// TIA Portal project "LaboratorioPID" (V21)

(* hardware
DEVICE "S7-1200 station_1"  S7-1200 Station
   slot 0: "Rack_0"  S7-1200 Rack  Rack  V1.0
   slot 1: "PLC-Serrato"  CPU 1214C AC/DC/Rly  6ES7 214-1BG40-0XB0  V4.2
   slot 3: "AQ 1x12BIT_1"  AQ1 signal board  6ES7 232-4HA30-0XB0  V1.0
DEVICE "HMI_1"  TP1200 Comfort
   slot 0: "HMI_1"  TP1200 Comfort  6AV2 124-0MC01-0AX0  17.0.0.0
   slot 1: "HMI_RT_1"  TP1200 Comfort  6AV2 124-0MC01-0AX0  17.0.0.0
   slot 5: "HMI_1.IE_CP_1"  PROFINET Interface  17.0.0.0
      slot 1: "PROFINET Interface_1"  PROFINET Interface
         slot 1: "Port_1"  Port
         slot 2: "Port_2"  Port
   slot 7: "HMI_1.MPI/DP_CP_1"  MPI/DP Interface  17.0.0.0
DEVICE "S7-1200 station_2"  S7-1200 Station
   slot 0: "Rack_0"  S7-1200 Rack  Rack  V1.0
   slot 1: "PLC-Liceth"  CPU 1214C AC/DC/Rly  6ES7 214-1BG40-0XB0  V4.2
*)

// ===== PLC "PLC-Serrato"  CPU 1214C AC/DC/Rly =====

VAR_GLOBAL   // PLC tag table "Default tag table"
   "PresionRaw" AT %IW64 : Int;
   "BelimoRaw" AT %QW80 : Int;
   "PID_salida_pct" AT %MD0 : Real;
   "Apertura_Manual" AT %MD10 : Real;
   "Clock_Byte" AT %MB100 : Byte;
   "Clock_10Hz" AT %M100.0 : Bool;
   "Clock_5Hz" AT %M100.1 : Bool;
   "Clock_2.5Hz" AT %M100.2 : Bool;
   "Clock_2Hz" AT %M100.3 : Bool;
   "Clock_1.25Hz" AT %M100.4 : Bool;
   "Clock_1Hz" AT %M100.5 : Bool;
   "Clock_0.625Hz" AT %M100.6 : Bool;
   "Clock_0.5Hz" AT %M100.7 : Bool;
   "PUT_DONE" AT %M20.0 : Bool;
   "PUT_ERROR" AT %M20.1 : Bool;
   "GET_NDR" AT %M20.2 : Bool;
   "GET_ERROR" AT %M20.3 : Bool;
   "PUT_STATUS" AT %MW22 : Word;
   "GET_STATUS" AT %MW24 : Word;
   "Tag_1" AT %MW20 : Word;
END_VAR

DATA_BLOCK "DBPresion"   // DB1
{ S7_Optimized_Access := 'TRUE' }
VERSION : 0.1
   VAR
      PresionBar : Real := 0.0;
      AperturaBelimo : Real := 0.0;
      AperturaManual : Real;
   END_VAR
BEGIN
END_DATA_BLOCK

DATA_BLOCK "DBHMI"   // DB2
{ S7_Optimized_Access := 'TRUE' }
VERSION : 0.1
   VAR
      Presión : Real;
      SP : Real;
      Modo : Bool;
      "Manual/Automatico" : Bool;
      PID_Manual : Bool;
   END_VAR
BEGIN
END_DATA_BLOCK

DATA_BLOCK "DBComunicacion"   // DB10
{ S7_Optimized_Access := 'FALSE' }
VERSION : 0.1
   VAR
      SP : Real;
      AperturaManual : Real;
      "Manual/Auto" : Bool;
      PresionBar : Real;
      AperturaBelimo : Real;
   END_VAR
BEGIN
END_DATA_BLOCK

FUNCTION "Vegabar_NS" : Void   // FC1, LAD
{ S7_Optimized_Access := 'TRUE' }
VERSION : 0.1
   VAR_TEMP
      PresionRaw : Int;
      PresionNorm : Real;
   END_VAR
BEGIN

REGION Network 1: Normalización y escalamiento de sensor
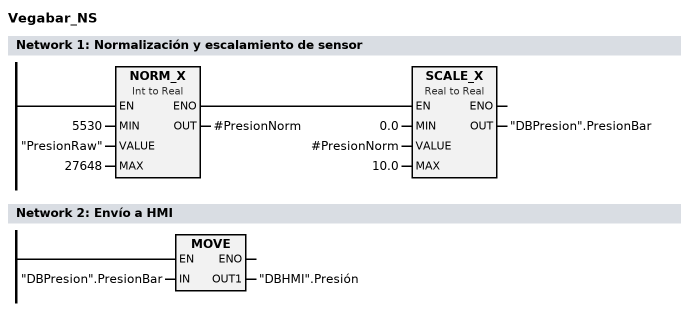
   RUNG wire#powerrail
      { S7_Templates := "[SrcType := Int, DestType := Real]" } Normalize(min := 5530, value := "PresionRaw", max := 27648, out => #PresionNorm)
      { S7_Templates := "[SrcType := Real, DestType := Real]" } Scale(min := 0.0, value := #PresionNorm, max := 10.0, out => "DBPresion".PresionBar)
   END_RUNG
   // the same network as SCL:
   #PresionNorm := NORM_X(MIN := 5530, VALUE := "PresionRaw", MAX := 27648);
   "DBPresion".PresionBar := SCALE_X(MIN := 0.0, VALUE := #PresionNorm, MAX := 10.0);
END_REGION

REGION Network 2: Envío a HMI
   RUNG wire#powerrail
      Move(in := "DBPresion".PresionBar, out1 => "DBHMI".Presión)
   END_RUNG
   // the same network as SCL:
   "DBHMI".Presión := "DBPresion".PresionBar;
END_REGION
END_FUNCTION

FUNCTION "Belimo_NS" : Void   // FC2, LAD
{ S7_Optimized_Access := 'TRUE' }
VERSION : 0.1
   VAR_TEMP
      BelimoNorm : Real;
   END_VAR
BEGIN

REGION Network 1: Modo manual
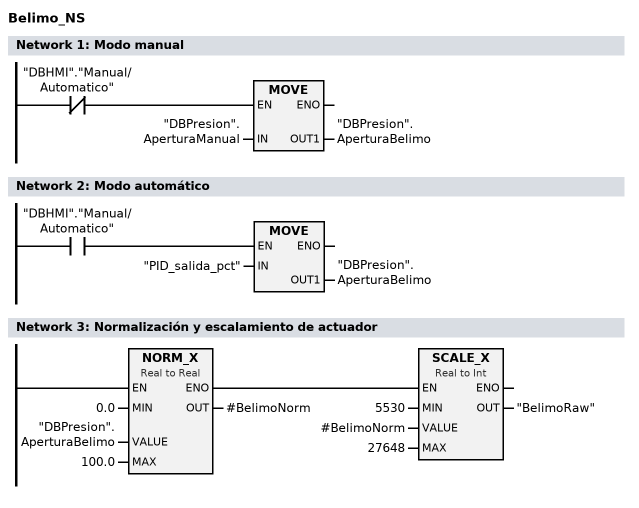
   RUNG wire#powerrail
      I_Contact( "DBHMI"."Manual/Automatico" )
      Move(in := "DBPresion".AperturaManual, out1 => "DBPresion".AperturaBelimo)
   END_RUNG
   // the same network as SCL:
   IF NOT "DBHMI"."Manual/Automatico" THEN "DBPresion".AperturaBelimo := "DBPresion".AperturaManual; END_IF;
END_REGION

REGION Network 2: Modo automático
   RUNG wire#powerrail
      Contact( "DBHMI"."Manual/Automatico" )
      Move(in := "PID_salida_pct", out1 => "DBPresion".AperturaBelimo)
   END_RUNG
   // the same network as SCL:
   IF "DBHMI"."Manual/Automatico" THEN "DBPresion".AperturaBelimo := "PID_salida_pct"; END_IF;
END_REGION

REGION Network 3: Normalización y escalamiento de actuador
   RUNG wire#powerrail
      { S7_Templates := "[SrcType := Real, DestType := Real]" } Normalize(min := 0.0, value := "DBPresion".AperturaBelimo, max := 100.0, out => #BelimoNorm)
      { S7_Templates := "[SrcType := Real, DestType := Int]" } Scale(min := 5530, value := #BelimoNorm, max := 27648, out => "BelimoRaw")
   END_RUNG
   // the same network as SCL:
   #BelimoNorm := NORM_X(MIN := 0.0, VALUE := "DBPresion".AperturaBelimo, MAX := 100.0);
   "BelimoRaw" := SCALE_X(MIN := 5530, VALUE := #BelimoNorm, MAX := 27648);
END_REGION
END_FUNCTION

FUNCTION "Comunicacion" : Void   // FC3, LAD
{ S7_Optimized_Access := 'TRUE' }
VERSION : 0.1
BEGIN

REGION Network 1: Bloque PUT
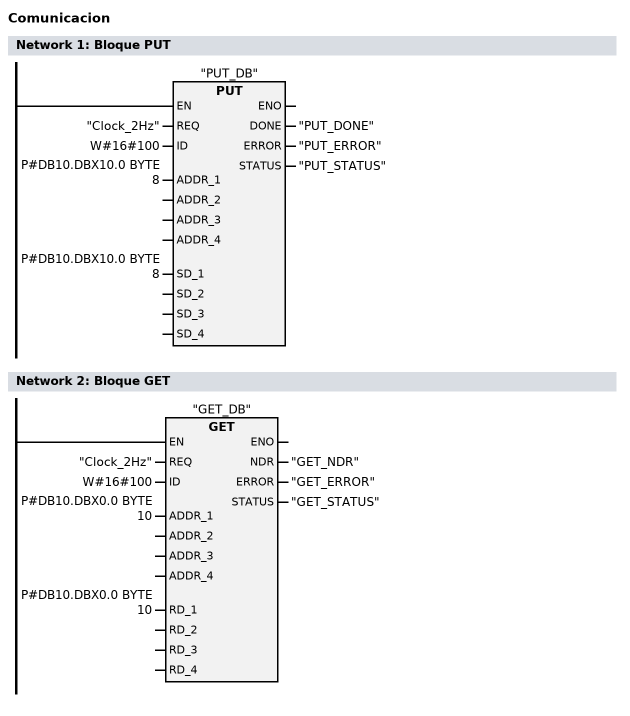
   "PUT_DB"(REQ := "Clock_2Hz",   // PUT
            ID := W#16#100,
            ADDR_1 := P#DB10.DBX10.0 BYTE 8,
            SD_1 := P#DB10.DBX10.0 BYTE 8,
            DONE => "PUT_DONE",
            ERROR => "PUT_ERROR",
            STATUS => "PUT_STATUS");
END_REGION

REGION Network 2: Bloque GET
   "GET_DB"(REQ := "Clock_2Hz",   // GET
            ID := W#16#100,
            ADDR_1 := P#DB10.DBX0.0 BYTE 10,
            RD_1 := P#DB10.DBX0.0 BYTE 10,
            NDR => "GET_NDR",
            ERROR => "GET_ERROR",
            STATUS => "GET_STATUS");
END_REGION
END_FUNCTION

ORGANIZATION_BLOCK "Main"   // OB1, LAD, ProgramCycle
TITLE = "Main Program Sweep (Cycle)"
{ S7_Optimized_Access := 'TRUE' }
VERSION : 0.1
   VAR_INPUT
      Initial_Call : Bool;   // Initial call of this OB
      Remanence : Bool;   // =True, if remanent data are available
   END_VAR
BEGIN

REGION Network 1: Bloque de sensor de presión
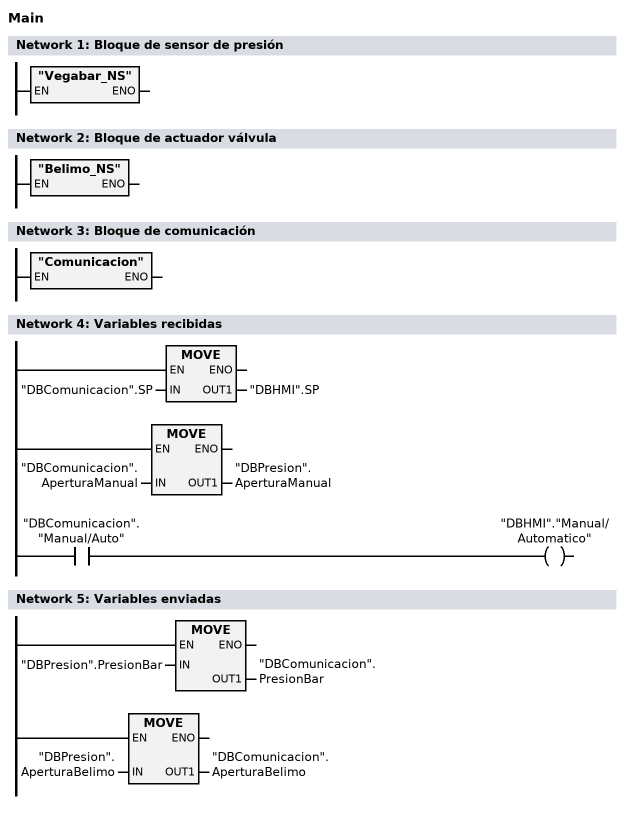
   RUNG wire#powerrail
      "Vegabar_NS"()
   END_RUNG
   // the same network as SCL:
   "Vegabar_NS"();
END_REGION

REGION Network 2: Bloque de actuador válvula
   RUNG wire#powerrail
      "Belimo_NS"()
   END_RUNG
   // the same network as SCL:
   "Belimo_NS"();
END_REGION

REGION Network 3: Bloque de comunicación
   RUNG wire#powerrail
      "Comunicacion"()
   END_RUNG
   // the same network as SCL:
   "Comunicacion"();
END_REGION

REGION Network 4: Variables recibidas
   RUNG wire#powerrail
      Move(in := "DBComunicacion".SP, out1 => "DBHMI".SP)
   END_RUNG
   RUNG wire#powerrail
      Move(in := "DBComunicacion".AperturaManual, out1 => "DBPresion".AperturaManual)
   END_RUNG
   RUNG wire#powerrail
      Contact( "DBComunicacion"."Manual/Auto" )
      Coil( "DBHMI"."Manual/Automatico" )
   END_RUNG
   // the same network as SCL:
   "DBHMI".SP := "DBComunicacion".SP;
   "DBPresion".AperturaManual := "DBComunicacion".AperturaManual;
   "DBHMI"."Manual/Automatico" := "DBComunicacion"."Manual/Auto";
END_REGION

REGION Network 5: Variables enviadas
   RUNG wire#powerrail
      Move(in := "DBPresion".PresionBar, out1 => "DBComunicacion".PresionBar)
   END_RUNG
   RUNG wire#powerrail
      Move(in := "DBPresion".AperturaBelimo, out1 => "DBComunicacion".AperturaBelimo)
   END_RUNG
   // the same network as SCL:
   "DBComunicacion".PresionBar := "DBPresion".PresionBar;
   "DBComunicacion".AperturaBelimo := "DBPresion".AperturaBelimo;
END_REGION
END_ORGANIZATION_BLOCK

ORGANIZATION_BLOCK "CyclicInterrupt"   // OB30, LAD, CyclicInterrupt
{ S7_Optimized_Access := 'TRUE' }
VERSION : 0.1
   VAR_INPUT
      Initial_Call : Bool;   // Initial call of this OB
      Event_Count : Int;   // Events discarded
   END_VAR
BEGIN

REGION Network 1: Habilitación de modo manual
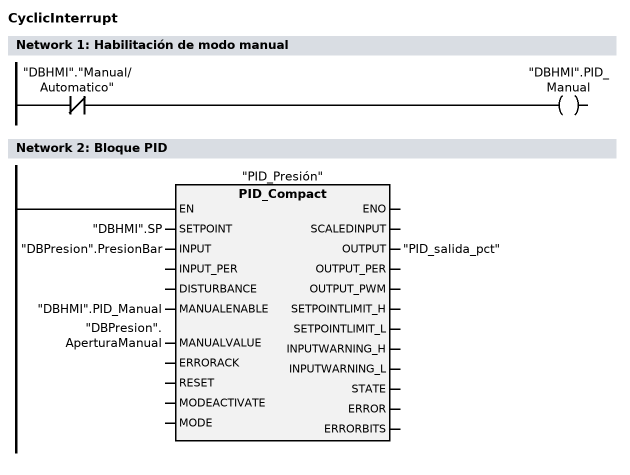
   RUNG wire#powerrail
      I_Contact( "DBHMI"."Manual/Automatico" )
      Coil( "DBHMI".PID_Manual )
   END_RUNG
   // the same network as SCL:
   "DBHMI".PID_Manual := NOT "DBHMI"."Manual/Automatico";
END_REGION

REGION Network 2: Bloque PID
   "PID_Presión"(Setpoint := "DBHMI".SP,   // PID_Compact
                 Input := "DBPresion".PresionBar,
                 ManualEnable := "DBHMI".PID_Manual,
                 ManualValue := "DBPresion".AperturaManual,
                 Output => "PID_salida_pct");
END_REGION
END_ORGANIZATION_BLOCK

// ===== PLC "PLC-Liceth"  CPU 1214C AC/DC/Rly =====

VAR_GLOBAL   // PLC tag table "Default tag table"
   "Clock_Byte" AT %MB100 : Byte;
   "Clock_10Hz" AT %M100.0 : Bool;
   "Clock_5Hz" AT %M100.1 : Bool;
   "Clock_2.5Hz" AT %M100.2 : Bool;
   "Clock_2Hz" AT %M100.3 : Bool;
   "Clock_1.25Hz" AT %M100.4 : Bool;
   "Clock_1Hz" AT %M100.5 : Bool;
   "Clock_0.625Hz" AT %M100.6 : Bool;
   "Clock_0.5Hz" AT %M100.7 : Bool;
   "PUT_DONE" AT %M20.0 : Bool;
   "PUT_ERROR" AT %M20.1 : Bool;
   "GET_NDR" AT %M20.2 : Bool;
   "GET_ERROR" AT %M20.3 : Bool;
   "PUT_STATUS" AT %MW22 : Word;
   "GET_STATUS" AT %MW24 : Word;
END_VAR

DATA_BLOCK "DBComunicacion"   // DB10
{ S7_Optimized_Access := 'FALSE' }
VERSION : 0.1
   VAR
      SP : Real;
      AperturaManual : Real;
      "Manual/Auto" : Bool;
      PresionBar : Real;
      AperturaBelimo : Real;
   END_VAR
BEGIN
END_DATA_BLOCK

FUNCTION "Comunicacion" : Void   // FC1, LAD
{ S7_Optimized_Access := 'TRUE' }
VERSION : 0.1
BEGIN

REGION Network 1: Bloque PUT
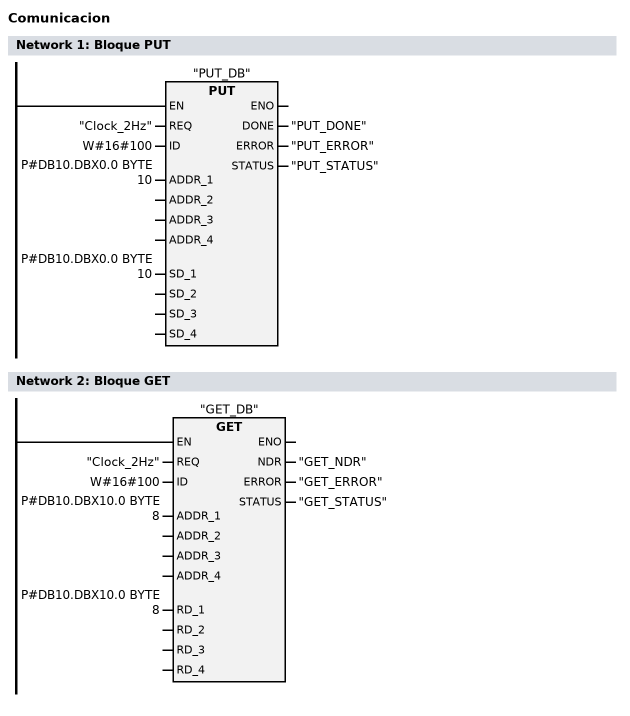
   "PUT_DB"(REQ := "Clock_2Hz",   // PUT
            ID := W#16#100,
            ADDR_1 := P#DB10.DBX0.0 BYTE 10,
            SD_1 := P#DB10.DBX0.0 BYTE 10,
            DONE => "PUT_DONE",
            ERROR => "PUT_ERROR",
            STATUS => "PUT_STATUS");
END_REGION

REGION Network 2: Bloque GET
   "GET_DB"(REQ := "Clock_2Hz",   // GET
            ID := W#16#100,
            ADDR_1 := P#DB10.DBX10.0 BYTE 8,
            RD_1 := P#DB10.DBX10.0 BYTE 8,
            NDR => "GET_NDR",
            ERROR => "GET_ERROR",
            STATUS => "GET_STATUS");
END_REGION
END_FUNCTION

ORGANIZATION_BLOCK "Main"   // OB1, LAD, ProgramCycle
TITLE = "Main Program Sweep (Cycle)"
{ S7_Optimized_Access := 'TRUE' }
VERSION : 0.1
   VAR_INPUT
      Initial_Call : Bool;   // Initial call of this OB
      Remanence : Bool;   // =True, if remanent data are available
   END_VAR
BEGIN

REGION Network 1: Bloque de comunicación
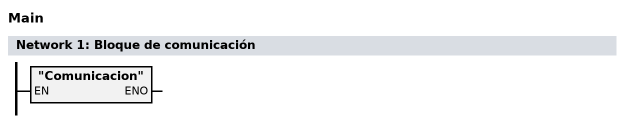
   RUNG wire#powerrail
      "Comunicacion"()
   END_RUNG
   // the same network as SCL:
   "Comunicacion"();
END_REGION
END_ORGANIZATION_BLOCK

(* ===== HMI "HMI_RT_1" =====
system functions are stored by id; their names below are inferred from use
connection "HMI_Connection_2": ETHERNET, S7_1200_OMS

HMI tags "Default tag table"
   "DBPresion_PresionBar" : Real = PLC DBComunicacion.PresionBar AT %DB10.DBD10, 1 s
   "DBHMI_SP" : Real = PLC DBComunicacion.SP AT %DB10.DBD0, 1 s
   "DBPresion_AperturaBelimo" : Real = PLC DBComunicacion.AperturaBelimo AT %DB10.DBD14, 1 s
   "DBHMI_Manual/Automatico" : Bool = PLC DBComunicacion.Manual/Auto AT %DB10.DBX8.0, 1 s
   "DBPresion_AperturaManual" : Real = PLC DBComunicacion.AperturaManual AT %DB10.DBD4, 1 s

screen "Root screen" 1280x800, template "Template_1"
   TextField "Text field_1" at 427,294 size 391x81; Text 'Laboratorio'
   TextField "Text field_2" at 243,382 size 788x81; Text 'PID de aire comprimido'
   GraphicView "Template_Graphic view_3" at 32,2 size 111x122; Picture "700863e0-019b-477d-b961-ae64ac70e2ac_1"

Template "Template_1" 1280x800
   Button "Exit" at 1200,739 size 78x59; TextOff 'Exit'; PictureOff "ExitRuntime_TP1200_Comfort_TR"; PictureOn "ExitRuntime_TP1200_Comfort_TR"
      on Release: StopRuntime(0)
   Button "Template_Button_11" at 241,739 size 78x59; TextOff 'AUTO'
      on Release: ActivateScreen("Auto", 0); SetBit("DBHMI_Manual/Automatico")
   Button "Alarms" at 81,739 size 78x59; TextOff 'Alarms'; PictureOff "AlarmDisplay_TP1200_Comfort_TR"; PictureOn "AlarmDisplay_TP1200_Comfort_TR"
      on Release: function_ef3f5d25("Alarm window_Unacknowledged", -1)
   Button "Start screen" at 1,739 size 78x59; TextOff 'Start screen'; PictureOff "NavigateHome_TP1200_Comfort_TR"; PictureOn "NavigateHome_TP1200_Comfort_TR"
      on Release: ActivateScreen("Root screen", 0)
   Button "Template_Button_12" at 161,739 size 78x59; TextOff 'MAN'
      on Release: ActivateScreen("Manual", 0); ResetBit("DBHMI_Manual/Automatico")

screen "Auto" 1280x800, template "Template_1"
   TextField "Text field_2" at 245,156 size 197x37; Text 'Presión (bar)'
   IOField "I/O field_1" at 246,242 size 206x89; FormatPattern 99.999
      ProcessValue <- "DBPresion_PresionBar"
   TextField "Text field_1" at 170,462 size 392x37; Text 'Apertura de la válvula (%)'
   IOField "I/O field_3" at 250,542 size 200x82; FormatPattern 999
      ProcessValue <- "DBPresion_AperturaBelimo"
   TextField "Text field_4" at 742,331 size 327x37; Text 'Setpoint presión (bar)'
   IOField "I/O field_2" at 784,408 size 219x107; FormatPattern 99.99
      ProcessValue <- "DBHMI_SP"
   TextField "Text field_3" at 416,29 size 445x62; Text 'Modo Automático'
   GraphicView "Template_Graphic view_3" at 32,2 size 111x122; Picture "700863e0-019b-477d-b961-ae64ac70e2ac_1"

screen "Manual" 1280x800, template "Template_1"
   TextField "Text field_2" at 277,330 size 197x37; Text 'Presión (bar)'
   IOField "I/O field_1" at 234,416 size 317x89; FormatPattern 99.9999999
      ProcessValue <- "DBPresion_PresionBar"
   TextField "Text field_1" at 693,331 size 392x37; Text 'Apertura de la válvula (%)'
   TextField "Text field_3" at 461,31 size 340x62; Text 'Modo Manual'
   GraphicView "Template_Graphic view_3" at 32,2 size 111x122; Picture "700863e0-019b-477d-b961-ae64ac70e2ac_1"
   IOField "I/O field_2" at 751,416 size 244x96; FormatPattern 999
      ProcessValue <- "DBPresion_AperturaManual"
*)